(* IEC 61131-3 sources: Twinova/app/src-tauri/project/tests/fixtures/valid/sort_line/components, 5 files *)

(* ---- twinova.belt@1.st ---- *)
(* Twinova belt conveyor, its drive, re-expressed from Open Industry Project's conveyor drive
   (examples/parts/_shared/conveyorDrive.js at 1e7488c, MIT). While the PLC's run is on, the surface ramps to
   speed_ref, which reads the speed parameter unless the PLC writes it: up at speed_at_30 per accel_time, down at
   speed_at_30 per decel_time, through 0 before it reverses; a ramp time of 0 is instant. running reports run after
   the start delay. The conveyor's native model reads surface_speed, and publishes the velocity, the encoder and the
   pulse itself. The field cycles every 1 ms, and TIME_TO_DWORD gives whole milliseconds, made a REAL through DINT:
   truST's DWORD_TO_REAL keeps the bits, not the number. n steps of speed_at_30 / n add up to speed_at_30 only within
   a rounding of REAL, so the ramp lands on its target within a hundredth of a step, on its millisecond. At its
   target the ramp is skipped. *)
FUNCTION_BLOCK BeltBehaviour
VAR_INPUT
    start_delay : TIME;
    accel_time : TIME;
    decel_time : TIME;
    speed_at_30 : REAL;
END_VAR
VAR_OUTPUT
    surface_speed : REAL;
END_VAR
VAR
    run AT %I* : BOOL;
    speed_ref AT %I* : REAL;
    running AT %Q* : BOOL;
    started : TON;
    target : REAL;
    ramp : TIME;
    step : REAL;
END_VAR
IF run THEN
    target := speed_ref;
ELSE
    target := 0.0;
END_IF;
IF target <> surface_speed THEN
    IF target * surface_speed < 0.0 THEN
        IF decel_time > T#0MS THEN
            target := 0.0;
        ELSE
            surface_speed := 0.0;
        END_IF;
    END_IF;
    IF ABS(target) > ABS(surface_speed) THEN
        ramp := accel_time;
    ELSE
        ramp := decel_time;
    END_IF;
    step := 0.0;
    IF ramp > T#0MS THEN
        step := speed_at_30 / DINT_TO_REAL(DWORD_TO_DINT(TIME_TO_DWORD(ramp)));
    END_IF;
    IF step <= 0.0 OR ABS(target - surface_speed) <= step * 1.01 THEN
        surface_speed := target;
    ELSIF target > surface_speed THEN
        surface_speed := surface_speed + step;
    ELSE
        surface_speed := surface_speed - step;
    END_IF;
END_IF;
started(IN := run, PT := start_delay);
running := started.Q;
END_FUNCTION_BLOCK

(* ---- twinova.pusher@1.st ---- *)
(* Twinova pusher, re-expressed from Open Industry Project's diverter (examples/parts/diverter/behavior.ts step() at
   1e7488c, MIT). extend sweeps the paddle out across its host; the reach slews linearly over push_time, out and back,
   as OIP's approach(). extended_fb and retracted_fb report the two ends of the stroke, which OIP shows only as its
   red and green lamps. The field cycles every 1 ms, so travel counts the milliseconds of stroke done, out of span. *)
FUNCTION_BLOCK PusherBehaviour
VAR_INPUT
    push_time : TIME;
END_VAR
VAR_OUTPUT
    reach : REAL;
END_VAR
VAR
    extend AT %I* : BOOL;
    extended_fb AT %Q* : BOOL;
    retracted_fb AT %Q* : BOOL;
    span : DINT;
    travel : DINT;
END_VAR
span := MAX(DWORD_TO_DINT(TIME_TO_DWORD(push_time)), 1);
IF extend THEN
    travel := MIN(travel + 1, span);
ELSE
    travel := MAX(travel - 1, 0);
END_IF;
reach := DINT_TO_REAL(travel) / DINT_TO_REAL(span);
extended_fb := travel = span;
retracted_fb := travel = 0;
END_FUNCTION_BLOCK

(* ---- twinova.roller@1.st ---- *)
(* Twinova roller conveyor, its drive, re-expressed from Open Industry Project's conveyor drive
   (examples/parts/_shared/conveyorDrive.js at 1e7488c, MIT). While the PLC's run is on, the surface ramps to
   speed_ref, which reads the speed parameter unless the PLC writes it: up at speed_at_30 per accel_time, down at
   speed_at_30 per decel_time, through 0 before it reverses; a ramp time of 0 is instant. running reports run after
   the start delay. The conveyor's native model reads surface_speed, and publishes the velocity, the encoder and the
   pulse itself. The field cycles every 1 ms, and TIME_TO_DWORD gives whole milliseconds, made a REAL through DINT:
   truST's DWORD_TO_REAL keeps the bits, not the number. n steps of speed_at_30 / n add up to speed_at_30 only within
   a rounding of REAL, so the ramp lands on its target within a hundredth of a step, on its millisecond. At its
   target the ramp is skipped. *)
FUNCTION_BLOCK RollerBehaviour
VAR_INPUT
    start_delay : TIME;
    accel_time : TIME;
    decel_time : TIME;
    speed_at_30 : REAL;
END_VAR
VAR_OUTPUT
    surface_speed : REAL;
END_VAR
VAR
    run AT %I* : BOOL;
    speed_ref AT %I* : REAL;
    running AT %Q* : BOOL;
    started : TON;
    target : REAL;
    ramp : TIME;
    step : REAL;
END_VAR
IF run THEN
    target := speed_ref;
ELSE
    target := 0.0;
END_IF;
IF target <> surface_speed THEN
    IF target * surface_speed < 0.0 THEN
        IF decel_time > T#0MS THEN
            target := 0.0;
        ELSE
            surface_speed := 0.0;
        END_IF;
    END_IF;
    IF ABS(target) > ABS(surface_speed) THEN
        ramp := accel_time;
    ELSE
        ramp := decel_time;
    END_IF;
    step := 0.0;
    IF ramp > T#0MS THEN
        step := speed_at_30 / DINT_TO_REAL(DWORD_TO_DINT(TIME_TO_DWORD(ramp)));
    END_IF;
    IF step <= 0.0 OR ABS(target - surface_speed) <= step * 1.01 THEN
        surface_speed := target;
    ELSIF target > surface_speed THEN
        surface_speed := surface_speed + step;
    ELSE
        surface_speed := surface_speed - step;
    END_IF;
END_IF;
started(IN := run, PT := start_delay);
running := started.Q;
END_FUNCTION_BLOCK

(* ---- twinova.stopper@1.st ---- *)
(* Twinova stopper, re-expressed from Open Industry Project's blade stop (examples/parts/blade-stop/part.js step()
   at 1e7488c, MIT). stop raises the blade; the lift slews linearly over raise_time, as OIP's approach() over its
   fixed 0.15 s. raised_fb reports the top of the stroke, which OIP does not have. The field cycles every 1 ms, so
   travel counts the milliseconds of stroke done; TIME_TO_DWORD gives whole milliseconds. *)
FUNCTION_BLOCK StopperBehaviour
VAR_INPUT
    raise_time : TIME;
END_VAR
VAR_OUTPUT
    lift : REAL;
END_VAR
VAR
    stop AT %I* : BOOL;
    raised_fb AT %Q* : BOOL;
    stroke : DINT;
    travel : DINT;
END_VAR
stroke := MAX(DWORD_TO_DINT(TIME_TO_DWORD(raise_time)), 1);
IF stop THEN
    travel := MIN(travel + 1, stroke);
ELSE
    travel := MAX(travel - 1, 0);
END_IF;
lift := DINT_TO_REAL(travel) / DINT_TO_REAL(stroke);
raised_fb := stop AND travel = stroke;
END_FUNCTION_BLOCK

(* ---- twinova.turntable@1.st ---- *)
(* Twinova turntable, re-expressed from Open Industry Project's turntable conveyor
   (examples/parts/turntable-conveyor/part.js step() at 1e7488c, MIT) and its conveyor drive
   (examples/parts/_shared/conveyorDrive.js). The deck slews the shortest way to target_angle, which reads the angle
   parameter unless the PLC writes it: up to rotation_speed over 0.5 s, braking to land on its target, and to a stop
   over 0.3 s while enable is off, resuming when it returns. Two changes from OIP: the deck starts at its angle
   parameter, not at 0, and a new target the other way ramps the turn through 0 instead of reversing it within a
   step. in_position reports the deck at rest on its target. The lane is a conveyor: while run is on and the deck is
   in position its surface ramps to speed_ref, as every conveyor's drive does (accel_time, decel_time, through 0
   before it reverses), and to 0 otherwise. The native model reads deck_angle (degrees, counter-clockwise seen from
   above), deck_rate (degrees per second) and surface_speed, and publishes the lane's velocity, encoder and pulse. The
   field cycles every 1 ms. *)
FUNCTION_BLOCK TurntableBehaviour
VAR_INPUT
    angle : REAL;
    rotation_speed : REAL;
    start_delay : TIME;
    accel_time : TIME;
    decel_time : TIME;
    speed_at_30 : REAL;
END_VAR
VAR_OUTPUT
    deck_angle : REAL;
    deck_rate : REAL;
    surface_speed : REAL;
END_VAR
VAR
    run AT %I* : BOOL;
    speed_ref AT %I* : REAL;
    target_angle AT %I* : REAL;
    enable AT %I* : BOOL;
    running AT %Q* : BOOL;
    in_position AT %Q* : BOOL;
    placed : BOOL;
    landed : BOOL;
    d : REAL;
    goal : REAL;
    change : REAL;
    started : TON;
    target : REAL;
    ramp : TIME;
    step : REAL;
END_VAR
IF NOT placed THEN
    deck_angle := angle;
    placed := TRUE;
END_IF;
d := target_angle - deck_angle;
IF d > 180.0 THEN
    d := d - 360.0;
ELSIF d <= -180.0 THEN
    d := d + 360.0;
END_IF;
change := rotation_speed / 0.5 * 0.001;
goal := 0.0;
IF NOT enable THEN
    change := rotation_speed / 0.3 * 0.001;
ELSIF deck_rate * d >= 0.0 AND ABS(d) > deck_rate * deck_rate / (rotation_speed / 0.5 * 2.0) THEN
    IF d > 0.0 THEN
        goal := rotation_speed;
    ELSE
        goal := -rotation_speed;
    END_IF;
END_IF;
IF deck_rate < goal THEN
    deck_rate := MIN(deck_rate + change, goal);
ELSE
    deck_rate := MAX(deck_rate - change, goal);
END_IF;
landed := deck_rate * d > 0.0 AND ABS(d) <= ABS(deck_rate) * 0.001;
IF landed THEN
    deck_angle := target_angle;
    deck_rate := 0.0;
ELSE
    deck_angle := deck_angle + deck_rate * 0.001;
END_IF;
IF deck_angle > 180.0 THEN
    deck_angle := deck_angle - 360.0;
ELSIF deck_angle <= -180.0 THEN
    deck_angle := deck_angle + 360.0;
END_IF;
in_position := deck_rate = 0.0 AND (landed OR d = 0.0);
IF run AND in_position THEN
    target := speed_ref;
ELSE
    target := 0.0;
END_IF;
IF target <> surface_speed THEN
    IF target * surface_speed < 0.0 THEN
        IF decel_time > T#0MS THEN
            target := 0.0;
        ELSE
            surface_speed := 0.0;
        END_IF;
    END_IF;
    IF ABS(target) > ABS(surface_speed) THEN
        ramp := accel_time;
    ELSE
        ramp := decel_time;
    END_IF;
    step := 0.0;
    IF ramp > T#0MS THEN
        step := speed_at_30 / DINT_TO_REAL(DWORD_TO_DINT(TIME_TO_DWORD(ramp)));
    END_IF;
    IF step <= 0.0 OR ABS(target - surface_speed) <= step * 1.01 THEN
        surface_speed := target;
    ELSIF target > surface_speed THEN
        surface_speed := surface_speed + step;
    ELSE
        surface_speed := surface_speed - step;
    END_IF;
END_IF;
started(IN := run, PT := start_delay);
running := started.Q;
END_FUNCTION_BLOCK
